(* IEC 61131-3 sources: trust-platform/examples/communication/ads_server_basic/src, 2 files *)

(* ---- config.st ---- *)
// The screens: after the task that calls Hmi.Display, the runtime copies the values they show,
// applies their commands and reads the alarms.
PROGRAM Screens
VAR
    Display : Hmi.Display;
END_VAR
    Display();
END_PROGRAM

CONFIGURATION Config
VAR_GLOBAL
    TankLevel : REAL := 42.5;
    PumpRunning : BOOL := FALSE;
    Setpoint : REAL := 10.0;
    StatusWord : WORD := 16#1234;
END_VAR
RESOURCE truST_ADS ON PLC
    TASK MainTask (INTERVAL := T#100ms, PRIORITY := 1);
    PROGRAM Main WITH MainTask : Main;
    TASK ScreenTask (INTERVAL := T#250ms, PRIORITY := 10);
    PROGRAM Screens WITH ScreenTask : Screens;
END_RESOURCE
END_CONFIGURATION

(* ---- main.st ---- *)
PROGRAM Main
VAR_EXTERNAL
    TankLevel : REAL;
    PumpRunning : BOOL;
    StatusWord : WORD;
END_VAR

// The program keeps TankLevel and PumpRunning moving. It leaves Setpoint, the writable
// symbol, to the ADS client, which reads back what it wrote.
TankLevel := TankLevel + 1.0;
IF TankLevel > 80.0 THEN
    TankLevel := 20.0;
END_IF;

PumpRunning := TankLevel > 40.0;
StatusWord := WORD#16#1234;
END_PROGRAM
